(* IEC 61131-3 sources: OpenPlc_Lezioni/conta_pezzi/build, 2 files *)

(* ---- plc.st ---- *)
TYPE
  LOGLEVEL : (CRITICAL, WARNING, INFO, DEBUG) := INFO;
END_TYPE

FUNCTION_BLOCK LOGGER
  VAR_INPUT
    TRIG : BOOL;
    MSG : STRING;
    LEVEL : LOGLEVEL := INFO;
  END_VAR
  VAR
    TRIG0 : BOOL;
  END_VAR

  IF TRIG AND NOT TRIG0 THEN
  {{
   LogMessage(GetFbVar(LEVEL),(char*)GetFbVar(MSG, .body),GetFbVar(MSG, .len));
  }}
  END_IF;
  TRIG0:=TRIG;
END_FUNCTION_BLOCK

PROGRAM program0
  VAR
    CTU0 : CTU;
    CU : BOOL;
    PULSE : BOOL;
    Q : BOOL;
    Reset : BOOL;
    Preset_value : INT := 5;
    R_TRIG1 : R_TRIG;
  END_VAR

  R_TRIG1(CLK := PULSE AND CU);
  CTU0(CU := R_TRIG1.Q, R := Reset, PV := Preset_value);
  Q := CTU0.Q;
END_PROGRAM

CONFIGURATION Config0

  RESOURCE Res0 ON PLC
    TASK task0(INTERVAL := T#20ms,PRIORITY := 0);
    PROGRAM instance0 WITH task0 : program0;
  END_RESOURCE
END_CONFIGURATION

(* ---- generated_plc.st ---- *)
PROGRAM program0
  VAR
    CTU0 : CTU;
    CU : BOOL;
    PULSE : BOOL;
    Q : BOOL;
    Reset : BOOL;
    Preset_value : INT := 5;
    R_TRIG1 : R_TRIG;
  END_VAR

  R_TRIG1(CLK := PULSE AND CU);
  CTU0(CU := R_TRIG1.Q, R := Reset, PV := Preset_value);
  Q := CTU0.Q;
END_PROGRAM

CONFIGURATION Config0

  RESOURCE Res0 ON PLC
    TASK task0(INTERVAL := T#20ms,PRIORITY := 0);
    PROGRAM instance0 WITH task0 : program0;
  END_RESOURCE
END_CONFIGURATION
